Fanuc KAREL source: KT00590.KL

PROGRAM KT00590
%NOLOCKGROUP
VAR
  S1: STRING[80]
  I2: INTEGER
  OUT: STRING[80]
BEGIN
  S1 = 'A'
    I2 = 3
  OUT = S1 + I2
END KT00590
